// TIA Portal V19 export
DATA_BLOCK "SPEED_COLD_SKID_CP02"   // DB109
// stored: InstanceOfName SPEED_REF_SCALING, InstanceOfType FB
"SPEED_REF_SCALING"
   // VAR_INPUT
   //    RAW_MIN : Int;
   //    RAW_MAX : Int;
   //    SCALE_MIN : Real;
   //    SCALE_MAX : Real;
   //    INPUT : Int;
   // END_VAR
   // VAR_OUTPUT
   //    SCALE_OUT : Int;
   // END_VAR
   // VAR
   //    SP : Real;
   // END_VAR
BEGIN
END_DATA_BLOCK
